(* IEC 61131-3 sources: trust-platform/examples/tutorials, 9 files *)

(* ---- 01_hello_counter.st ---- *)
PROGRAM HelloCounter
VAR
    enable : BOOL := TRUE;
    reset_cmd : BOOL := FALSE;
    increment : DINT := 1;
    count : DINT := 0;
END_VAR

IF reset_cmd THEN
    count := 0;
ELSIF enable THEN
    count := count + increment;
END_IF;
END_PROGRAM

(* ---- 02_blinker.st ---- *)
PROGRAM Blinker
VAR
    enable : BOOL := TRUE;
    lamp : BOOL := FALSE;
    pulse_pt : TIME := T#250ms;
    timer_enable : BOOL := TRUE;
    blink_timer : TON;
END_VAR

blink_timer(IN := timer_enable, PT := pulse_pt);

IF NOT enable THEN
    lamp := FALSE;
    timer_enable := FALSE;
ELSIF blink_timer.Q THEN
    lamp := NOT lamp;
    timer_enable := FALSE;
ELSE
    timer_enable := TRUE;
END_IF;
END_PROGRAM

(* ---- 03_traffic_light.st ---- *)
PROGRAM TrafficLight
VAR
    phase : INT := 0;
    phase_pt : TIME := T#500ms;
    phase_timer_enable : BOOL := TRUE;
    phase_timer : TON;
    red : BOOL := TRUE;
    yellow : BOOL := FALSE;
    green : BOOL := FALSE;
END_VAR

phase_timer(IN := phase_timer_enable, PT := phase_pt);

CASE phase OF
    0:
        red := TRUE;
        yellow := FALSE;
        green := FALSE;
    1:
        red := TRUE;
        yellow := TRUE;
        green := FALSE;
    2:
        red := FALSE;
        yellow := FALSE;
        green := TRUE;
    3:
        red := FALSE;
        yellow := TRUE;
        green := FALSE;
END_CASE;

IF phase_timer.Q THEN
    CASE phase OF
        0:
            phase := 1;
        1:
            phase := 2;
        2:
            phase := 3;
        3:
            phase := 0;
    END_CASE;
    phase_timer_enable := FALSE;
ELSE
    phase_timer_enable := TRUE;
END_IF;
END_PROGRAM

(* ---- 04_tank_level.st ---- *)
PROGRAM TankLevel
VAR
    inlet_valve_cmd : BOOL := FALSE;
    outlet_valve_cmd : BOOL := TRUE;
    level_percent : REAL := 45.0;
    low_setpoint : REAL := 30.0;
    high_setpoint : REAL := 70.0;
END_VAR

IF level_percent <= low_setpoint THEN
    inlet_valve_cmd := TRUE;
    outlet_valve_cmd := FALSE;
ELSIF level_percent >= high_setpoint THEN
    inlet_valve_cmd := FALSE;
    outlet_valve_cmd := TRUE;
END_IF;

IF inlet_valve_cmd THEN
    level_percent := level_percent + 2.5;
END_IF;

IF outlet_valve_cmd THEN
    level_percent := level_percent - 1.5;
END_IF;
END_PROGRAM

(* ---- 05_motor_starter.st ---- *)
PROGRAM MotorStarter
VAR
    start_pb : BOOL := FALSE;
    stop_pb : BOOL := FALSE;
    overload_trip : BOOL := FALSE;
    motor_run : BOOL := FALSE;
    seal_in_contact : BOOL := FALSE;
END_VAR

IF stop_pb OR overload_trip THEN
    motor_run := FALSE;
ELSIF start_pb OR seal_in_contact THEN
    motor_run := TRUE;
END_IF;

seal_in_contact := motor_run;
END_PROGRAM

(* ---- 06_recipe_manager.st ---- *)
PROGRAM RecipeManager
VAR
    selected_recipe : INT := 1;
    apply_selection : BOOL := TRUE;
    active_target_temp : REAL := 0.0;
    active_mix_time : TIME := T#0s;
    active_batch_size : INT := 0;
END_VAR

IF apply_selection THEN
    CASE selected_recipe OF
        1:
            active_target_temp := 65.0;
            active_mix_time := T#30s;
            active_batch_size := 10;
        2:
            active_target_temp := 72.5;
            active_mix_time := T#45s;
            active_batch_size := 14;
        3:
            active_target_temp := 80.0;
            active_mix_time := T#60s;
            active_batch_size := 18;
        ELSE
            active_target_temp := 60.0;
            active_mix_time := T#20s;
            active_batch_size := 8;
    END_CASE;
END_IF;
END_PROGRAM

(* ---- 07_pid_loop.st ---- *)
PROGRAM PidLoop
VAR
    setpoint : REAL := 50.0;
    process_value : REAL := 40.0;
    kp : REAL := 1.2;
    ki : REAL := 0.1;
    kd : REAL := 0.05;
    sample_time : REAL := 0.1;
    integral_term : REAL := 0.0;
    previous_error : REAL := 0.0;
    error : REAL := 0.0;
    derivative : REAL := 0.0;
    control_output : REAL := 0.0;
END_VAR

error := setpoint - process_value;
integral_term := integral_term + (error * ki * sample_time);
derivative := (error - previous_error) / sample_time;
control_output := (kp * error) + integral_term + (kd * derivative);
previous_error := error;
process_value := process_value + (control_output * 0.02);
END_PROGRAM

(* ---- 08_conveyor_system.st ---- *)
PROGRAM ConveyorSystem
VAR
    start_cmd : BOOL := FALSE;
    stop_cmd : BOOL := FALSE;
    jam_sensor : BOOL := FALSE;
    part_at_entry : BOOL := FALSE;
    part_at_exit : BOOL := FALSE;
    conveyor_run : BOOL := FALSE;
    reject_gate : BOOL := FALSE;
    part_counter : DINT := 0;
END_VAR

IF stop_cmd OR jam_sensor THEN
    conveyor_run := FALSE;
ELSIF start_cmd THEN
    conveyor_run := TRUE;
END_IF;

IF conveyor_run AND part_at_entry THEN
    reject_gate := FALSE;
END_IF;

IF conveyor_run AND part_at_exit THEN
    part_counter := part_counter + 1;
END_IF;

IF jam_sensor THEN
    reject_gate := TRUE;
END_IF;
END_PROGRAM

(* ---- 09_simulation_coupling.st ---- *)
PROGRAM SimulationCouplingDemo
VAR
    tank_level_raw : WORD;
    high_level_alarm : BOOL;
END_VAR

high_level_alarm := WORD_TO_UINT(tank_level_raw) >= 500;
END_PROGRAM

CONFIGURATION SimulationCouplingConfig
TASK Cycle (INTERVAL := T#100ms, PRIORITY := 1);
PROGRAM P1 WITH Cycle : SimulationCouplingDemo;
VAR_CONFIG
    P1.tank_level_raw AT %IW0 : WORD;
    P1.high_level_alarm AT %QX0.0 : BOOL;
END_VAR
END_CONFIGURATION
